Staubli VAL3: V20201012.pgx

program V20201012()
begin
  //Version: V1.2
  //Date: February 14, 2020
  //Editor: Zhang Huajun
  //  1.Improved real-time position display, can view joints and Cartesian coordinates
  //  2.Improve popup information display
  //  3.Corrected the error that the target point cannot be reached

  //Version: V1.3
  //Date: April 9, 2020
  //Editor: Zhang Huajun
  //  1.Reduce unnecessary binding
  //  2.Use CSS to keep Stäubli SP2 interface style
  //
  //
  //Version: V2.0
  //Date: August 20, 2020
  //Editor: Zhang Huajun
  //  1.Optimize HMI response by turning libsave() into a background task
  //  2.Optimize widgets binding
  //
  //
  //Version: V2.1
  //Date: October 12, 2020
  //Editor: Zhang Huajun
  //  1.Add 2 points to calculate TCP for 4-axis robot (only output X and Y)
end
